// TIA Portal V21 export
// export: Created 2026-10-23T20:43:04.5564133Z, ExportSetting WithDefaults, DisplayName Totally Integrated Automation Portal, DisplayVersion V21 Update 1, DisplayName SINAMICS Startdrive Advanced, DisplayVersion V21 HF2, DisplayName SINAMICS Startdrive G110M, G120, G120C, G120D, G120P, G115D, DisplayVersion V21 HF2, DisplayName SINAMICS Startdrive G130, G150, S120, S150, G200, G220, S200, S210, S220, Innomotics MVD, DisplayVersion V21 HF2, DisplayName STEP 7 Professional, DisplayVersion V21 Update 1, DisplayName STEP 7 Safety, DisplayVersion V21, DisplayName Tech WebApplication, DisplayVersion V21, DisplayName WinCC Basic/Comfort/Advanced, DisplayVersion V21 Update 1, DisplayName WinCC Unified, DisplayVersion V21 Update 1
DATA_BLOCK "IDB_FbdBoxes"   // DB22
VERSION : 0.1
// stored: AutoNumber true, DBAccessibleFromOPCUA true, DBAccessibleFromWebserver true, InstanceOfName FB_FbdBoxes, InstanceOfType FB
"FB_FbdBoxes"
   // VAR_INPUT
   //    Start : Bool;
   //    InValue : Int;
   //    Limit : Int;
   // END_VAR
   // VAR_OUTPUT
   //    Delayed : Bool;
   //    Copy : Int;
   //    Sum : Int;
   //    IsEqual : Bool;
   //    SectionsOk : Bool;
   //    Skipped : Bool;
   //    AfterJump : Bool;
   // END_VAR
   // VAR
   //    Delay { S7_SetPoint := 'True'} : TON_TIME;
   //    DelayElapsed : Time;
   //    Timers { S7_SetPoint := 'True'} : "FB_SclTimers";
   //    TimerRunOn : Bool;
   //    TimerPulse : Bool;
   //    TimerCount : Int;
   //    TimerDelayed : Bool;
   //    TimerReached : Bool;
   // END_VAR
BEGIN
END_DATA_BLOCK
